Yaskawa INFORM job: MAINCAL.JBI

/JOB
//NAME MAINCAL
//POS
///NPOS 1,0,1,0,0,0
///TOOL 9
///POSTYPE PULSE
///PULSE
C00000=0,0,0
EC00000=0
//INST
<volatile>
///COMM Generated using RoboDK
///ATTR SC,RW
///GROUP1 RB1
NOP
'Program generated by RoboDK v
'6.0.7 for Yaskawa Motoman EPL
'160 on XX/XX/XXXX 18:00:00
'Using nominal kinematics.
'Using Frame S (targets wrt ba
'se):
'1234.6,-98.8,50.5,0.0,0.0,30.
'0
MOVJ C00000 VJ=50.00  +MOVJ EC00000 VJ=100.00
CALL JOB:SUBPROG
CALL JOB:NOTAPRO
END
